(* IEC 61131-3 sources: llm-plc-st-eval/data/raw/claude-sonnet-4-6/B2/zero_shot, 3 files *)

(* ---- ejec_1.st ---- *)
```pascal
FUNCTION_BLOCK FB_Valvula
VAR_INPUT
    nivelAlto : BOOL; (* Sensor de nivel alto del tanque *)
END_VAR

VAR_OUTPUT
    valvula : BOOL; (* TRUE = válvula abierta, FALSE = válvula cerrada *)
END_VAR

VAR
    tonRetardo : TON; (* Temporizador on-delay de 5 segundos *)
END_VAR

(* -------------------------------------------------------
   Lógica de control:
   - El temporizador se habilita solo mientras nivelAlto
     esté activo de forma continua.
   - Si nivelAlto cae a FALSE, el temporizador se resetea
     inmediatamente (IN := FALSE) y la válvula cierra.
   - Cuando el temporizador completa T#5S (Q = TRUE),
     la válvula abre.
   ------------------------------------------------------- *)

(* Llamada al temporizador: se activa con nivelAlto *)
tonRetardo(
    IN := nivelAlto,   (* Habilita el conteo mientras nivel esté alto *)
    PT := T#5S         (* Tiempo de retardo requerido *)
);

(* La válvula abre cuando el temporizador completa los 5 s.
   Si nivelAlto cae, tonRetardo.Q vuelve FALSE de inmediato
   porque IN := FALSE resetea el bloque TON. *)
valvula := tonRetardo.Q;

END_FUNCTION_BLOCK
```

(* ---- ejec_2.st ---- *)
```pascal
FUNCTION_BLOCK FB_Valvula
VAR_INPUT
    nivelAlto : BOOL; (* Sensor de nivel alto del tanque *)
END_VAR

VAR_OUTPUT
    valvula : BOOL; (* TRUE = válvula abierta, FALSE = válvula cerrada *)
END_VAR

VAR
    tonRetardo : TON; (* Temporizador on-delay para confirmar nivel alto *)
END_VAR

(* ---------------------------------------------------------------
   Lógica de control:
   - El temporizador TON se habilita mientras nivelAlto esté activo.
   - Si nivelAlto permanece TRUE durante 5 s continuos, tonRetardo.Q
     se pone TRUE y la válvula abre.
   - Si nivelAlto cae a FALSE en cualquier momento, el temporizador
     se resetea (IN=FALSE) y la válvula cierra de inmediato.
--------------------------------------------------------------- *)

(* Llamada al temporizador: se activa solo si nivelAlto es TRUE *)
tonRetardo(
    IN  := nivelAlto,
    PT  := T#5S
);

(* La válvula abre cuando el temporizador confirma 5 s de nivel alto;
   cierra de inmediato si nivelAlto deja de estar activo *)
valvula := tonRetardo.Q;

END_FUNCTION_BLOCK
```

(* ---- ejec_3.st ---- *)
```pascal
FUNCTION_BLOCK FB_Valvula
VAR_INPUT
    nivelAlto : BOOL; (* Sensor de nivel alto del tanque *)
END_VAR

VAR_OUTPUT
    valvula : BOOL; (* TRUE = válvula abierta, FALSE = válvula cerrada *)
END_VAR

VAR
    tonRetardo : TON; (* Temporizador on-delay para confirmar nivel alto *)
END_VAR

(* ---------------------------------------------------------------
   Lógica de control:
   - El temporizador TON se habilita mientras nivelAlto esté activo.
   - Si nivelAlto permanece TRUE durante 5 s continuos, tonRetardo.Q
     se pone TRUE y abre la válvula.
   - Si nivelAlto cae a FALSE en cualquier momento, el temporizador
     se resetea (IN=FALSE) y la válvula cierra de inmediato.
--------------------------------------------------------------- *)

(* Llamada al temporizador: se activa con nivelAlto, tiempo de 5 s *)
tonRetardo(
    IN := nivelAlto,
    PT := T#5S
);

(* La válvula abre solo cuando el temporizador ha completado los 5 s *)
valvula := tonRetardo.Q;

END_FUNCTION_BLOCK
```
